(* IEC 61131-3 sources: lasal-git-demo/CPU/LasalDemoProject/Network, 1 file *)

(* ---- ConfigObjects.st ---- *)
FUNCTION GLOBAL TAB TASK_CONF
_K_TASK, _K_REAL,
_K_END_VAR,

_K_TASK, _K_CYCLIC,
_K_END_VAR,

_K_TASK, _K_BACKGROUND,
_K_END_VAR,

_K_END_CONF
END_FUNCTION

FUNCTION GLOBAL TAB IPR_CONF
_K_IPR
	0$UINT,
_K_END_VAR,
_K_END_CONF
END_FUNCTION

FUNCTION GLOBAL TAB CONFIG_TABLES
00089$UINT,
0$UINT, 1, 15, "_BUSINTERFACESDIASDRIVEMNG",
0$UINT, 0, 5, "_CAN",
0$UINT, 1, 11, "_CANLIB",
0$UINT, 1, 72, "_DRIVEAXIS",
0$UINT, 1, 81, "_DRIVEAXISBASE",
0$UINT, 1, 22, "_DRIVEAXISSET",
0$UINT, 1, 88, "_DRIVEMNG_DC061",
0$UINT, 1, 88, "_DRIVEMNG_DC101",
0$UINT, 1, 66, "_DRIVEMNGBASE",
0$UINT, 1, 20, "_FILESYS",
0$UINT, 0, 5, "_LINKER",
0$UINT, 1, 1, "_MULTITASK",
0$UINT, 1, 9, "_OPENSSL",
0$UINT, 0, 5, "_OSKERNEL",
0$UINT, 1, 36, "_SERLIB",
0$UINT, 2, 0, "_STDLIB",
0$UINT, 1, 3, "_SYNCMEASURE",
0$UINT, 1, 2, "_SYNCMEASUREECAT",
0$UINT, 0, 0, "_SYSMSG",
0$UINT, 1, 1, "_TASKOBJECTCONTROL",
0$UINT, 1, 6, "_USERLOGGING",
0$UINT, 1, 69, "_VARANDRIVEBASE",
0$UINT, 1, 21, "ASCII_BIN",
0$UINT, 1, 26, "BUSINTERFACESDIAS",
0$UINT, 2, 1, "BUSINTERFACESDIASINTERNAL",
0$UINT, 1, 1, "CP112_IOS",
0$UINT, 1, 0, "CP313_IOS",
0$UINT, 0, 4, "CRITICALSECTION",
0$UINT, 0, 0, "DEMOCLASS",
0$UINT, 1, 42, "DI200",
0$UINT, 2, 33, "DIASMASTER",
0$UINT, 1, 83, "DIASMASTERC",
0$UINT, 2, 25, "DIASMASTERMAIN",
0$UINT, 1, 0, "DIASMASTERPOSTSCAN",
0$UINT, 2, 2, "ECAT_MASTER_BASE",
0$UINT, 2, 0, "ECAT_SLAVE_BASE",
0$UINT, 1, 11, "EEPROM",
0$UINT, 1, 0, "ENVBASE",
0$UINT, 1, 1, "ENVIRONMENTVARIABLE",
0$UINT, 1, 0, "ENVLIB",
0$UINT, 1, 0, "ENVSTRINGACTION",
0$UINT, 1, 1, "ETHERCAT_HUB_BASE",
0$UINT, 2, 2, "ETHERCAT_PLC",
0$UINT, 1, 4, "GETCILINTERFACE",
0$UINT, 1, 21, "HUB_BASE",
0$UINT, 2, 11, "HUB_BASE_ROOT",
0$UINT, 2, 36, "HWBASE",
0$UINT, 2, 56, "HWBASECDIAS",
0$UINT, 1, 0, "HWCLOGGING",
0$UINT, 5, 27, "HWCONTROL",
0$UINT, 1, 10, "HWCONTROLBASE",
0$UINT, 1, 0, "HWRTPOSTSCAN",
0$UINT, 1, 6, "I2CCDIAS",
0$UINT, 1, 22, "MERKEREX",
0$UINT, 7, 2, "OPC_UA",
0$UINT, 2, 0, "OPC_UA_BASE",
0$UINT, 1, 0, "OPC_UA_DATALOGGERBASE",
0$UINT, 1, 0, "OPC_UA_ENCRYPTIONBASE",
0$UINT, 1, 1, "OPC_UA_INTERFACE",
0$UINT, 1, 7, "OPC_UA_MODULEBASE",
0$UINT, 1, 0, "OPC_UA_OPENSSL_V1_1_1",
0$UINT, 3, 0, "OPC_UA_SERVER",
0$UINT, 1, 17, "RAMEX",
0$UINT, 1, 9, "RAMFILE",
0$UINT, 1, 39, "SAFETYBASEFSOE",
0$UINT, 3, 19, "SAFETYCDIAS_BASE",
0$UINT, 2, 30, "SAFETYMANAGER",
0$UINT, 1, 4, "SAFETYUDP",
0$UINT, 1, 11, "SCP211",
0$UINT, 1, 23, "SDI101",
0$UINT, 1, 60, "SDIASBASE",
0$UINT, 1, 10, "SDIASHUBBASE",
0$UINT, 1, 99, "SDIASMANAGER",
0$UINT, 2, 8, "SDIASPLC",
0$UINT, 1, 10, "SDIASSAFETYBASE",
0$UINT, 1, 41, "SDIASSAFETYMANAGERFSOE",
0$UINT, 0, 46, "SIGCLIB",
0$UINT, 1, 23, "STO081",
0$UINT, 1, 11, "STRING",
0$UINT, 1, 86, "STRINGINTERNAL",
0$UINT, 1, 21, "SYNCCALL",
0$UINT, 1, 34, "TO161",
0$UINT, 2, 21, "VARAN_BASE",
0$UINT, 3, 8, "VARANMANAGER",
0$UINT, 2, 8, "VARANMANAGER_1",
0$UINT, 1, 26, "VARANMANAGER_BASE",
0$UINT, 1, 3, "VIRTUALBASEINIT",
0$UINT, 2, 11, "WATCHDOGDIAS",
0$UINT, 1, 2, "XXXBASE_IOS",
ONE_CFG$UINT, 0, 0, "ONE_DemoNetwork",
ONE_CFG$UINT, 0, 0, "ONE_HW_Network",
TASK_CFG$UINT, 0, 0, "TASK_CONF",
IPR_CFG$UINT, 0, 0, "IPR_CONF",
PRJ_CFG$UINT, 0, 0, "LasalDemoProject",
END_FUNCTION

FUNCTION GLOBAL TAB CH_REDIRECT_EMB_TAB
0000$UINT,
00033$UINT,
"_BUSINTERFACESDIASDRIVEMNG;SERIALNO", "\SERIALNOSTR.DATA",
"_DRIVEMNG_DC061;FWDATETR", "\FWDATESTRING.DATA",
"_DRIVEMNG_DC061;FWDATE", "\FWDATESTRING.DATA",
"_DRIVEMNG_DC061;FWNUMSTR", "\FWNUMSTRING.DATA",
"_DRIVEMNG_DC061;FWVERSION", "\FWNUMSTRING.DATA",
"_DRIVEMNG_DC101;FWDATETR", "\FWDATESTRING.DATA",
"_DRIVEMNG_DC101;FWDATE", "\FWDATESTRING.DATA",
"_DRIVEMNG_DC101;FWNUMSTR", "\FWNUMSTRING.DATA",
"_DRIVEMNG_DC101;FWVERSION", "\FWNUMSTRING.DATA",
"_USERLOGGING;ENV_EVENTLOGLEVELNAME", "\ENVVAR_FORWLVL\ENVNAME.DATA",
"_USERLOGGING;ENV_FILELOGLEVELNAME", "\ENVVAR_LOGLVL\ENVNAME.DATA",
"_VARANDRIVEBASE;SERIALNO", "\SERIALNOSTR.DATA",
"BUSINTERFACESDIAS;SERIALNO", "\SERIALNOSTR.DATA",
"DI200;SERIALNO", "\SERIALNOSTR.DATA",
"ECAT_MASTER_BASE;SOFTWAREVERSION", "\STRSOFTWAREVERSION.DATA",
"ECAT_SLAVE_BASE;DEVICENAME", "\DEVICENAMESTR.DATA",
"ECAT_SLAVE_BASE;PRODUCTREVISION", "\PRODUCTREVSTR.DATA",
"ENVIRONMENTVARIABLE;SSTRINGVALUE", "\ENVVALUE.DATA",
"ENVIRONMENTVARIABLE;SVARIABLENAME", "\ENVNAME.DATA",
"ETHERCAT_PLC;SOFTWAREVERSION", "\STRSOFTWAREVERSION.DATA",
"HWBASECDIAS;SERIALNO", "\SERIALNOSTR.DATA",
"SAFETYCDIAS_BASE;SERIALNO", "\SERIALNOSTR.DATA",
"SCP211;DESIGNERPRJNAME", "\SDIASSAFETYMANAGERFSOE1\PROJECTNAMESTR.DATA",
"SCP211;DESIGNERPRJREV", "\SDIASSAFETYMANAGERFSOE1\PROJECTREVISIONSTR.DATA",
"SCP211;SERIALNO", "\SERIALNOSTR.DATA",
"SDI101;SERIALNO", "\SERIALNOSTR.DATA",
"SDIASBASE;SERIALNO", "\SERIALNOSTR.DATA",
"SDIASSAFETYBASE;SERIALNO", "\SERIALNOSTR.DATA",
"SDIASSAFETYMANAGERFSOE;DESIGNERPRJNAME", "\PROJECTNAMESTR.DATA",
"SDIASSAFETYMANAGERFSOE;DESIGNERPRJREV", "\PROJECTREVISIONSTR.DATA",
"STO081;SERIALNO", "\SERIALNOSTR.DATA",
"TO161;SERIALNO", "\SERIALNOSTR.DATA",
"VARAN_BASE;SERIALNO", "\SERIALNOSTR.DATA",
END_FUNCTION
